FUNCTION_BLOCK ArmCartesian
VAR
    stage : INT;
    i : INT;
    k : INT;
    curve : ARRAY[0..16] OF LREAL;
    incoming : ARRAY[0..16] OF LREAL;
    p : ARRAY[1..5] OF LREAL;
    v : ARRAY[1..5] OF LREAL;
    a : ARRAY[1..5] OF LREAL;
    dir : ARRAY[1..5] OF DINT;
    velocity_limit : ARRAY[1..5] OF LREAL;
    acceleration_limit : ARRAY[1..5] OF LREAL;
    deceleration_limit : ARRAY[1..5] OF LREAL;
    jerk_limit : ARRAY[1..5] OF LREAL;
    elapsed : LREAL;
    phase_elapsed : LREAL;
    cycle_seconds : LREAL;
    segment_seconds : LREAL;
    u : LREAL;
    path_progress : LREAL;
    ds : LREAL;
    dds : LREAL;
    delta : LREAL;
    bend : LREAL;
    slope_bound : LREAL;
    allowed : BOOL;
    drive_ready : BOOL;
    all_enabled : BOOL;
    all_disabled : BOOL;
    all_stopped : BOOL;
    all_released : BOOL;
    arrived : BOOL;
    reject_error : UDINT;
    last_heartbeat : UDINT;
    heartbeat_age : LREAL;
    finish_state : UDINT;
    fb_enable : ARRAY[1..5] OF MC_ExtSetPointGenEnable;
    fb_disable : ARRAY[1..5] OF MC_ExtSetPointGenDisable;
    fb_stop : ARRAY[1..5] OF MC_Stop;
END_VAR

// 定位臂归零保留原1ms曲线接口，第16项必须为0。
cycle_seconds := UDINT_TO_LREAL(TwinCAT_SystemInfoVarList._TaskInfo[1].CycleTime) * 0.0000001;
IF TwinCAT_SystemInfoVarList._TaskInfo[1].FirstCycle THEN
    G.arm_curve_ack := G.arm_curve_request;
    G.arm_curve_cancel := TRUE;
    G.arm_curve_owned := FALSE;
    G.arm_curve_state := 0;
    G.arm_curve_error := 0;
    stage := 0;
END_IF
IF G.arm_curve_heartbeat <> last_heartbeat THEN
    last_heartbeat := G.arm_curve_heartbeat;
    heartbeat_age := 0;
ELSE
    heartbeat_age := heartbeat_age + cycle_seconds;
END_IF

drive_ready := G.arm_manual_enable AND NOT G.host_comm_timeout AND NOT G.estop_hold_req
    AND (ABS(cycle_seconds - 0.001) < 0.00000001);
FOR i := 1 TO 5 DO
    drive_ready := drive_ready AND G.arm_power_output[i].Done AND G.arm_enable_req[i]
        AND NOT G.arm_axis[i].Status.Error AND NOT G.arm_reset_req[i]
        AND NOT G.arm_jog_pos_req[i] AND NOT G.arm_jog_neg_req[i];
END_FOR
allowed := drive_ready AND (heartbeat_age < 0.5);

IF G.arm_curve_request <> G.arm_curve_ack THEN
    IF stage >= 40 THEN
        // 停止中的迟到请求只确认接收，不重新启动运动。
        IF G.arm_curve_error = 0 THEN G.arm_curve_error := 2001; END_IF
        finish_state := 4;
        G.arm_curve_cancel := TRUE;
        G.arm_curve_ack := G.arm_curve_request;
    ELSE
        reject_error := 0;
        FOR k := 0 TO 16 DO
            incoming[k] := G.arm_curve_data[k];
            IF NOT ((incoming[k] >= -100000.0) AND (incoming[k] <= 100000.0)) THEN
                reject_error := 2002;
            END_IF
        END_FOR
        IF (incoming[15] < 0.02) OR (incoming[15] > 120.0)
            OR (incoming[16] <> 0.0) THEN
            reject_error := 2002;
        END_IF
        IF NOT allowed OR G.arm_curve_cancel THEN reject_error := 2003; END_IF
        IF (stage <> 0) AND (reject_error = 0) THEN reject_error := 2001; END_IF
        IF G.arm_cjog_owned THEN reject_error := 2001; END_IF

        IF reject_error = 0 THEN
            FOR i := 1 TO 5 DO
                IF NOT ((G.arm_jog_velocity[i] > 0) AND (G.arm_jog_velocity[i] <= 10000))
                    OR NOT ((G.arm_jog_acc[i] > 0) AND (G.arm_jog_acc[i] <= 10000))
                    OR NOT ((G.arm_jog_dec[i] > 0) AND (G.arm_jog_dec[i] <= 10000))
                    OR NOT ((G.arm_jog_jerk[i] > 0) AND (G.arm_jog_jerk[i] <= 10000)) THEN
                    reject_error := 2002;
                END_IF
            END_FOR
        END_IF
        IF reject_error = 0 THEN
            FOR i := 1 TO 5 DO
                delta := incoming[i+4] - incoming[i-1];
                segment_seconds := incoming[15];
                    bend := incoming[i+9];
                    IF ABS(bend) > ABS(delta)/4.0+0.000000001 THEN reject_error := 2002; END_IF
                    slope_bound := ABS(delta)+4.0*ABS(bend);
                    IF (1.875*slope_bound/segment_seconds > G.arm_jog_velocity[i]+0.0000001)
                        OR ((6.0*slope_bound+28.125*ABS(bend))/(segment_seconds*segment_seconds)
                            > G.arm_jog_acc[i]+0.0000001) THEN
                        reject_error := 2005;
                    END_IF

            END_FOR
            IF (MIN(incoming[4],incoming[9]) < -60.0)
                OR (MAX(incoming[4],incoming[9]) > 60.0) THEN reject_error := 2006; END_IF
        END_IF
        IF reject_error = 0 THEN
            FOR i := 1 TO 5 DO
                // 负载下反馈会波动，启动只依据忙状态，不用速度或起点偏差判停稳。
                IF G.arm_motion_busy[i] THEN
                    reject_error := 2004;
                END_IF
            END_FOR
        END_IF

        IF reject_error = 0 THEN
                FOR k := 0 TO 16 DO curve[k] := incoming[k]; END_FOR
                FOR i := 1 TO 5 DO
                    p[i] := curve[i-1];
                    v[i] := 0;
                    a[i] := 0;
                    dir[i] := 0;
                    IF curve[i+4] > p[i] THEN dir[i] := 1; END_IF
                    IF curve[i+4] < p[i] THEN dir[i] := -1; END_IF
                    velocity_limit[i] := G.arm_jog_velocity[i];
                    acceleration_limit[i] := G.arm_jog_acc[i];
                    deceleration_limit[i] := G.arm_jog_dec[i];
                    jerk_limit[i] := G.arm_jog_jerk[i];
                END_FOR
                G.arm_curve_owned := TRUE;
                stage := 10;
                elapsed := 0;
                phase_elapsed := 0;
                finish_state := 2;
                G.arm_curve_progress := 0;
            G.arm_curve_error := 0;
            G.arm_curve_state := 1;
        ELSE
            IF G.arm_curve_error = 0 THEN G.arm_curve_error := reject_error; END_IF
            G.arm_curve_cancel := TRUE;
            finish_state := 4;
            IF stage > 0 THEN
                stage := 40;
                phase_elapsed := 0;
            END_IF
        END_IF
        // 先锁存归零曲线，再确认序号。
        G.arm_curve_ack := G.arm_curve_request;
    END_IF
END_IF

IF (stage > 0) AND (stage < 40) THEN
    IF G.arm_curve_cancel OR NOT allowed THEN
        finish_state := 3;
        IF NOT allowed THEN
            IF G.arm_curve_error = 0 THEN G.arm_curve_error := 2003; END_IF
            finish_state := 4; G.arm_curve_cancel := TRUE;
        END_IF
        stage := 40;
        phase_elapsed := 0;
    END_IF
END_IF
IF stage > 0 THEN phase_elapsed := phase_elapsed + cycle_seconds; END_IF
IF (stage = 10 OR stage = 30) AND (phase_elapsed > 2.0) THEN
    IF G.arm_curve_error = 0 THEN G.arm_curve_error := 2007; END_IF
    G.arm_curve_cancel := TRUE;
    finish_state := 4;
    stage := 40;
END_IF

IF stage = 20 THEN
    u := MIN(1.0, elapsed/curve[15]);
    path_progress := u*u*u*(10.0+u*(-15.0+6.0*u));
    ds := 30.0*u*u*(1.0-u)*(1.0-u)/curve[15];
    dds := 60.0*u*(1.0-u)*(1.0-2.0*u)/(curve[15]*curve[15]);
    FOR i := 1 TO 5 DO
        delta := curve[i+4]-curve[i-1];
            bend := curve[i+9];
            p[i] := curve[i-1]+path_progress*delta+4.0*path_progress*(1.0-path_progress)*bend;
            v[i] := (delta+4.0*(1.0-2.0*path_progress)*bend)*ds;
            a[i] := (delta+4.0*(1.0-2.0*path_progress)*bend)*dds-8.0*bend*ds*ds;
        IF (ABS(v[i]) > velocity_limit[i]+0.000001)
            OR (ABS(a[i]) > acceleration_limit[i]+0.000001)
            OR NOT ((G.arm_act_pos[i]-p[i] >= -1.0) AND (G.arm_act_pos[i]-p[i] <= 1.0)) THEN
            IF G.arm_curve_error = 0 THEN G.arm_curve_error := 2008; END_IF
            G.arm_curve_cancel := TRUE;
            finish_state := 4;
            stage := 40;
        END_IF
    END_FOR
    G.arm_curve_progress := u;
    elapsed := elapsed+cycle_seconds;
    IF (u >= 1.0) AND (stage = 20) THEN
        stage := 30;
        phase_elapsed := 0;
    END_IF
END_IF

all_enabled := TRUE;
all_disabled := TRUE;
all_stopped := TRUE;
all_released := TRUE;
arrived := TRUE;
FOR i := 1 TO 5 DO
    // 归零沿用原外部设定点发生器握手。
    IF G.arm_curve_owned THEN
        MC_ExtSetPointGenFeed(Axis:=G.arm_axis[i], Position:=p[i],
            Velocity:=v[i], Acceleration:=a[i], Direction:=dir[i]);
    END_IF
    fb_enable[i](Axis:=G.arm_axis[i], Execute:=(stage=10),
        Position:=curve[i+4], PositionType:=POSITIONTYPE_ABSOLUTE);
    fb_disable[i](Axis:=G.arm_axis[i], Execute:=(stage=40));
    fb_stop[i](Axis:=G.arm_axis[i], Execute:=(stage=50) AND NOT G.arm_axis[i].Status.Error,
        Deceleration:=deceleration_limit[i], Jerk:=jerk_limit[i]);
    all_enabled := all_enabled AND fb_enable[i].Enabled;
    // 与末端点动相同，错误轴和功能块错误不阻塞所有权释放。
    all_disabled := all_disabled AND (fb_disable[i].Done OR fb_disable[i].Error OR G.arm_axis[i].Status.Error);
    all_stopped := all_stopped AND (fb_stop[i].Done OR fb_stop[i].Error OR G.arm_axis[i].Status.Error);
    all_released := all_released AND NOT fb_stop[i].Busy;
    arrived := arrived AND (ABS(G.arm_act_pos[i]-curve[i+4]) <= 0.05)
        AND (ABS(G.arm_act_vel[i]) <= 0.1);
    IF G.arm_curve_owned AND (fb_enable[i].Error OR fb_disable[i].Error OR fb_stop[i].Error) THEN
        G.arm_curve_cancel := TRUE;
        IF G.arm_curve_error = 0 THEN
            IF fb_enable[i].Error THEN G.arm_curve_error := fb_enable[i].ErrorID;
            ELSIF fb_disable[i].Error THEN G.arm_curve_error := fb_disable[i].ErrorID;
            ELSIF fb_stop[i].Error THEN G.arm_curve_error := fb_stop[i].ErrorID; END_IF
        END_IF
        finish_state := 4;
        IF stage < 40 THEN stage := 40; END_IF
    END_IF
END_FOR

CASE stage OF
10:
    IF all_enabled THEN stage := 20; elapsed := 0; phase_elapsed := 0; END_IF
30:
    IF arrived AND (phase_elapsed >= 2.0*cycle_seconds) THEN stage := 40; END_IF
40:
    IF all_disabled THEN
        IF finish_state = 2 THEN stage := 60; ELSE stage := 50; END_IF
    END_IF
50:
    IF all_stopped THEN stage := 60; END_IF
60:
    IF all_released THEN
        G.arm_curve_owned := FALSE;
        G.arm_curve_state := finish_state;
        stage := 0;
    END_IF
END_CASE
IF G.arm_curve_error <> 0 THEN
    G.arm_curve_state := 4;
END_IF

END_FUNCTION_BLOCK

(* stored: Version 1.1.0.1, ProductVersion 3.1.4024.15
   POU ArmCartesian: Id {713355bc-7855-44d6-b270-717a93d9e329}, SpecialFunc None *)
